(* IEC 61131-3 sources: plc-st-test/packages/cli/test/fixtures/failing/src, 1 file *)

(* ---- FB_Counter.st ---- *)
FUNCTION_BLOCK FB_Counter
VAR_INPUT
  bEnable : BOOL;
END_VAR
VAR_OUTPUT
  nCount : DINT;
END_VAR
IF bEnable THEN
  nCount := nCount + 1;
END_IF
END_FUNCTION_BLOCK
